// TIA Portal V17 export
FUNCTION "FC_T01_Contacts" : Void   // FC101, LAD
{ S7_Optimized_Access := 'TRUE' }
// stored: SetENOAutomatically false
   VAR_INPUT
      Marche : Bool;
      Arret : Bool;
      Capteur_A : Bool;
      Capteur_B : Bool;
   END_VAR
   VAR_OUTPUT
      Sortie_Serie : Bool;
   END_VAR
   VAR_IN_OUT
      Moteur : Bool;
   END_VAR
BEGIN

REGION Network 1: Auto-maintien marche / arrêt
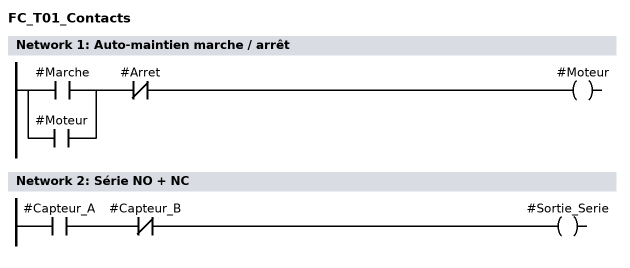
   RUNG wire#powerrail
      Contact( #Marche )
      wire#w1
      I_Contact( #Arret )
      Coil( #Moteur )
   END_RUNG
   RUNG wire#powerrail
      Contact( #Moteur )
   END_RUNG wire#w1
   // the same network as SCL:
   #Moteur := (#Marche OR #Moteur) AND NOT #Arret;
END_REGION

REGION Network 2: Série NO + NC
   RUNG wire#powerrail
      Contact( #Capteur_A )
      I_Contact( #Capteur_B )
      Coil( #Sortie_Serie )
   END_RUNG
   // the same network as SCL:
   #Sortie_Serie := #Capteur_A AND NOT #Capteur_B;
END_REGION
END_FUNCTION
